// TIA Portal V20 export
// export: Created 2026-10-20T12:45:40.5766009Z, ExportSetting WithDefaults, DisplayName Totally Integrated Automation Portal, DisplayVersion V20 Update 6, DisplayName TIA Portal Openness, DisplayVersion V20 Update 6, DisplayName TIA Portal Version Control Interface, DisplayVersion V20 Update 6, DisplayName SINAMICS Startdrive Advanced, DisplayVersion V20 SP1, DisplayName SINAMICS Startdrive G130, G150, S120, S150, SINAMICS MV, G220, S200, S210, DisplayVersion V20 SP1, DisplayName SINAMICS Startdrive G110M, G120, G120C, G120D, G120P, G115D, DisplayVersion V20 SP1, DisplayName STEP 7 Professional, DisplayVersion V20 Update 6, DisplayName STEP 7 Safety, DisplayVersion V20 Update 2, DisplayName WinCC Basic/Comfort/Advanced, DisplayVersion V20 Update 6, DisplayName WinCC Unified, DisplayVersion V20 Update 6
DATA_BLOCK "HMI_OrderTable"   // DB110
{ S7_Optimized_Access := 'TRUE' }
VERSION : 0.1
// stored: AutoNumber true, DBAccessibleFromOPCUA true, IsOnlyStoredInLoadMemory false, IsRetainMemResEnabled false, IsWriteProtectedInAS false, MemoryReserve 100
   VAR
      OrderTable : Array[0..9] of "OrderTable_UDT";
      State { S7_SetPoint := 'True'} : Array[0..9] of USInt;
      Index : Array[0..9] of Int;
      ScrollUp_PB : Bool;
      ScrollDown_PB : Bool;
      PlaceOrder_PB : Bool;
      PauseOrders_PB : Bool;
      ResumeOrder_PB : Bool;
      CancelOrder_PB : Bool;
      CancelThisOrder_PB : Bool;
      StartRow : Int;
      Device : USInt;
      PlacingNewOrder : Bool;
      PopUp_ErrorWindow_Active : Bool;
      PopUp_ErrorID : UInt;
      PopUp_Index : Int;
   END_VAR
BEGIN
END_DATA_BLOCK
